(* IEC 61131-3 sources: Codesys_IAP/Demo/PLC1/Magazijn Overzetter Simulatie Structured Text 2V1 - Leeg_tekst/Programma Structured Text/StationClass, 8 files *)

(* ---- cycle.st ---- *)
(*#### DECLARATIE ####*)
// Datum : 26 november 2026, Auteur: Gerard Harkema
METHOD cycle
VAR
END_VAR
(*#### IMPLEMENTATIE ####*)
// TODO: implementeer volgens het statediagram van StationClass

(* ---- initialize.st ---- *)
(*#### DECLARATIE ####*)
// Datum : 26 november 2026, Auteur: Gerard Harkema
METHOD initialize
VAR_INPUT
	IORef			: REFERENCE TO stationIO;
END_VAR
(*#### IMPLEMENTATIE ####*)
IO REF= IORef;

// Elk object krijgt zijn eigen IO-structuur
magazijn.initialize(IO.magazijn);
overzetter.initialize(IO.overzetter);

eState := stationStates.idle;

(* ---- isError.st ---- *)
(*#### DECLARATIE ####*)
// Datum : 26 november 2026, Auteur: Gerard Harkema
METHOD isError : BOOL
VAR_INPUT
END_VAR
(*#### IMPLEMENTATIE ####*)
// TODO: implementeer volgens het statediagram van StationClass

(* ---- isKlaar.st ---- *)
(*#### DECLARATIE ####*)
// Datum : 26 november 2026, Auteur: Gerard Harkema
METHOD isKlaar : BOOL
VAR_INPUT
END_VAR
(*#### IMPLEMENTATIE ####*)
// TODO: implementeer volgens het statediagram van StationClass

(* ---- isMagazijnLeeg.st ---- *)
(*#### DECLARATIE ####*)
// Datum : 26 november 2026, Auteur: Gerard Harkema
METHOD isMagazijnLeeg : BOOL
VAR_INPUT
END_VAR
(*#### IMPLEMENTATIE ####*)
// TODO: implementeer volgens het statediagram van StationClass

(* ---- noodstop.st ---- *)
(*#### DECLARATIE ####*)
// Datum : 26 november 2026, Auteur: Gerard Harkema
METHOD noodstop
VAR_INPUT
END_VAR
(*#### IMPLEMENTATIE ####*)
// TODO: implementeer volgens het statediagram van StationClass

(* ---- reset.st ---- *)
(*#### DECLARATIE ####*)
// Datum : 26 november 2026, Auteur: Gerard Harkema
METHOD reset
VAR_INPUT
END_VAR
(*#### IMPLEMENTATIE ####*)
// TODO: implementeer volgens het statediagram van StationClass

(* ---- start.st ---- *)
(*#### DECLARATIE ####*)
// Datum : 26 november 2026, Auteur: Gerard Harkema
METHOD start : BOOL
VAR_INPUT
END_VAR
(*#### IMPLEMENTATIE ####*)
// TODO: implementeer volgens het statediagram van StationClass
